Staubli VAL3: physicalIO.pgx

program physicalIO()
// TX60 Level 1 IO adapter: bIn2 cylinder presence; valve1 gripper.
begin
  // ============================================================
  // E/S DEL TX60: PINZA AJUSTADA AL MANDO MANUAL T1
  // ============================================================
  // start solo crea esta tarea si simulation=false al arrancar.
  // Una lectura DIO necesita comparacion: bIn2 == true devuelve bool.
  // No usar directamente wait(io:bIn2), que da "invalid type".
  //
  // bIn0: sensor de presencia en herramienta para buscar pistones
  //        en Level 3. NO es confirmacion de pieza agarrada.
  // bOut10: extender/retraer el alimentador de cilindros, Level 2.
  // bIn14/bIn15: finales extendido/retraido de ese alimentador.
  // Estas cuatro senales no intervienen en nuestro Level 1.
  while true
    // bIn2=1: hay cilindro preparado; bIn2=0: no detecta cilindro.
    cylinderPresent = io:bIn2 == true

    // El enunciado indicaba bOut0; en esta celda T1 usa valve1.
    // El usuario confirma que la pinza responde al mando manual.
    // valve1=1 ABRE; valve1=0 CIERRA. No copiar la logica de vacio de 2A.
    // Una sola pinza para tLateral y tTip; el adaptador solo lee presencia.
    // TODO FISICO: comprobar respuesta real antes del primer recorrido.
    // La pinza se manda desde start con open/close; no sobrescribir valve1.

    // Primera lectura/escritura realizada; start ya puede continuar.
    ioReady = true
    delay(0.01)
  endWhile
end
